Fanuc KAREL source: KA00058.KL

PROGRAM KA00058
%NOLOCKGROUP
VAR
  SRC: POSITION
  DST: CONFIG
BEGIN
  DST = SRC
END KA00058
